(* IEC 61131-3 sources: s7-to-codesys/src/POUs/Lang/Converted/FC_ClampPctLad, 2 files *)

(* ---- FC_ClampPctLad.decl.st ---- *)
// Назначение: Ограничение значения пределами (LAD)
//             Результат: iIn, ограниченный снизу iMin и сверху iMax (сначала верхний предел, затем нижний). ENO не
//             пишется: ENO = EN.
// Автор:      WTP2 (исходный блок S7); перевод в ST — s7conv 0.1.0
// Версия:     0.1 (исходный блок S7)
// Документ:   docs/CONVERSION_REPORT.md, docs/MAPPING.md
// Источник:   samples/lang/FC_ClampPctLad.xml, LAD, SW.Blocks.FC "FC_ClampPctLad", пространство имён Interface/v5,
//             FAMILY Utils
// Сгенерировано s7conv: пометки MIGRATION-CHECK и MIGRATION-TODO требуют ручного разбора.
FUNCTION FC_ClampPctLad : INT
VAR_INPUT
    iIn : INT;  // Значение
    iMin : INT;  // Нижний предел
    iMax : INT;  // Верхний предел
END_VAR

(* ---- FC_ClampPctLad.impl.st ---- *)
// Сеть 1: Значение по умолчанию
FC_ClampPctLad := iIn;
// Сеть 2: Выше максимума
IF iIn > iMax THEN
    FC_ClampPctLad := iMax;
END_IF
// Сеть 3: Ниже минимума
IF iIn < iMin THEN
    FC_ClampPctLad := iMin;
END_IF
